// TwinCAT 3 PLC project Untitled1
// ProgramVersion: 3.1.4026.25
// libraries:
//   Tc2_Standard, * (Beckhoff Automation GmbH)
//   Tc2_System, * (Beckhoff Automation GmbH)
// project tree:
//   GVLs/ GVL_EverySignal.TcGVL, GVL_Inputs.TcGVL, GVL_IO.TcGVL, GVL_Outputs.TcGVL
//   / PlcTask.TcTTO
//   POUs/ MAIN.TcPOU, PRG_Mapping.TcPOU
// real-time tasks:
//   TASK PlcTask: cycle T#10ms, priority 20, ADS port 350
//   TASK PlcTask1: cycle T#10ms, priority 21, ADS port 351
//   TASK CNC-Task ADS: cycle default, priority 7, ADS port 558
//   TASK CNC-Task COM: cycle T#10ms, priority 14, ADS port 556
//   TASK CNC-Task SDA: cycle T#10ms, priority 9, ADS port 555
//   TASK CNC-Task GEO: cycle T#2ms, priority 3, ADS port 554
// motion (NC):
//   TASK NC-Task 1 SAF: cycle T#2ms, priority 4, ADS port 501
//   TASK NC-Task 1 SVB: cycle T#10ms, priority 8, ADS port 511
//   AXIS Axis 1 (id 1)
//     OtherSettings: AllowMotionCmdToSlave=true
//     encoder EncType=8
//       EncPara: MaxCount=#xffffffff
//     drive DrvType=9
//       DrvPara: MaxCount=#xffffffff
//         Analog: VeloScale=6, TorqueSetpointScale=10, ScaleFactorActTorque=0.1
//         TimeComp: TaskDelayCycles=1
//     controller CtrType=1
//       CtrPara: PriorControlFactor=1
//         Observer: BandWidth=20
//   AXIS Axis 2 (id 2)
//     OtherSettings: AllowMotionCmdToSlave=true
//     encoder EncType=8
//       EncPara: MaxCount=#xffffffff
//     drive DrvType=9
//       DrvPara: MaxCount=#xffffffff
//         Analog: VeloScale=6, TorqueSetpointScale=10, ScaleFactorActTorque=0.1
//         TimeComp: TaskDelayCycles=1
//     controller CtrType=1
//       CtrPara: PriorControlFactor=1
//         Observer: BandWidth=20
// I/O:
//   DEVICE C6015 (X102), AmsNetId 192.168.0.101.2.1
//     EtherCAT1  (CU1128) Junction [CU1128 6x EtherCAT junction] // Connected to PLC (C6015) using X1
//       (AX5206-0000-0011) EtherCAT4 [AX5206-0000-0011 EtherCAT Drive (SoE, 2 Ch.)] // Attached to EtherCAT1 at EtherCAT
//       EtherCAT2  (EK1100) Coupler MP-6K1 [EK1100 EtherCAT Coupler (2A E-Bus)] // Connected to EtherCAT1, Junction at X1 (W EtherCAT2 RS PRO 240-6302 1m 4x0.14 5.1)
//         (EL1809) Input Terminal MP-6K10 [EL1809 16Ch. Dig. Input 24V, 3ms] // Attached to EtherCAT 2 Coupler
//         (EL2809) Output Teminal MP-6K20 [EL2809 16Ch. Dig. Output 24V, 0.5A] // Attached to EtherCAT2 Coupler
//       Box 8 (EP1018-0001) MS-9K1 [EP1018-0001 8 Ch. Dig. Input 24V, 10µs, M8]
//       Box 9 (EP1018-0001) MS-9K2 [EP1018-0001 8 Ch. Dig. Input 24V, 10µs, M8]
//       Box 10 (EP1018-0001) MS-9K3 [EP1018-0001 8 Ch. Dig. Input 24V, 10µs, M8]
//       Box 11 (EP2028-0001) MS-10K1 [EP2028-0001 8 Ch. Dig. Output 24V, 2A, M8]
//       Box 12 (EP2028-0001) MS-10K2 [EP2028-0001 8 Ch. Dig. Output 24V, 2A, M8]
//       EtherCAT3 (EK1100) Coupler LS-7K1 [EK1100 EtherCAT Coupler (2A E-Bus)] // Attached to EtherCAT1, Junction at X1 (W EtherCAT3 RS PRO 240-6325 5m 4x0.14)
//         (EL1809) Input Terminal LS-7K10 [EL1809 16Ch. Dig. Input 24V, 3ms] // Attached to EtherCAT3 Coupler
//         (EL2809) Output Terminal LS-7K20 [EL2809 16Ch. Dig. Output 24V, 0.5A] // Attached to EtherCAT3 Coupler
//       Box 2 (CU1128-B) [CU1128 6x EtherCAT junction - Dev A]
//       Box 3 (CU1128-C) [CU1128 6x EtherCAT junction - Dev B]
// variable links:
//   Untitled1/Untitled1 Instance <-> C6015 (X102)/EtherCAT1  (CU1128) Junction/Box 10 (EP1018-0001) MS-9K3
//     PlcTask Inputs/GVL_IO.DI_E1052_{0..7} <-> Channel {1..8}/E1052.{0..7}_X{1..8}:4_DI{0..7}  (8 links)
//   Untitled1/Untitled1 Instance <-> C6015 (X102)/EtherCAT1  (CU1128) Junction/Box 11 (EP2028-0001) MS-10K1
//     PlcTask Outputs/GVL_IO.DQ_A1050_{0..7} <-> Channel {1..8}/A1050.{0..7}_X{1..8}:4_DQ{0..7}  (8 links)
//   Untitled1/Untitled1 Instance <-> C6015 (X102)/EtherCAT1  (CU1128) Junction/Box 12 (EP2028-0001) MS-10K2
//     PlcTask Outputs/GVL_IO.DQ_A1051_{0..7} <-> Channel {1..8}/A1051.{0..7}_X{1..8}:4_DQ{0..7}  (8 links)
//   Untitled1/Untitled1 Instance <-> C6015 (X102)/EtherCAT1  (CU1128) Junction/Box 8 (EP1018-0001) MS-9K1
//     PlcTask Inputs/GVL_IO.DI_E1050_0 <-> Channel 1/E1050.0 _X1:4_DI0
//     PlcTask Inputs/GVL_IO.DI_E1050_{1..5} <-> Channel {2..6}/E1050.{1..5}_X{2..6}:4_DI{1..5}  (5 links)
//   Untitled1/Untitled1 Instance <-> C6015 (X102)/EtherCAT1  (CU1128) Junction/Box 9 (EP1018-0001) MS-9K2
//     PlcTask Inputs/GVL_IO.DI_E1051_{0..3} <-> Channel {1..4}/E1051.{0..3}_X{1..4}:4_DI{0..3}  (4 links)
//   Untitled1/Untitled1 Instance <-> C6015 (X102)/EtherCAT1  (CU1128) Junction/EtherCAT2  (EK1100) Coupler MP-6K1/(EL1809) Input Terminal MP-6K10
//     PlcTask Inputs/GVL_IO.DI_E0_0 <-> Channel 1/E0.0_1_DI0
//     PlcTask Inputs/GVL_IO.DI_E0_1 <-> Channel 2/E0.1_2_DI1
//   Untitled1/Untitled1 Instance <-> C6015 (X102)/EtherCAT1  (CU1128) Junction/EtherCAT2  (EK1100) Coupler MP-6K1/(EL2809) Output Teminal MP-6K20
//     PlcTask Outputs/GVL_IO.DQ_A0_0 <-> Channel 1/A0.0_1_DQ0
//     PlcTask Outputs/GVL_IO.DQ_A0_1 <-> Channel 2/A0.1_2_DQ1
//   Untitled1/Untitled1 Instance <-> C6015 (X102)/EtherCAT1  (CU1128) Junction/EtherCAT3 (EK1100) Coupler LS-7K1/ (EL2809) Output Terminal LS-7K20
//     PlcTask Outputs/GVL_IO.DQ_A50_{0..5} <-> Channel {1..6}/A50.{0..5}_{1..6}_DQ{0..5}  (6 links)
//   Untitled1/Untitled1 Instance <-> C6015 (X102)/EtherCAT1  (CU1128) Junction/EtherCAT3 (EK1100) Coupler LS-7K1/(EL1809) Input Terminal LS-7K10
//     PlcTask Inputs/GVL_IO.DI_E50_0 <-> Channel 1/E50.0_1_DI0
//     PlcTask Inputs/GVL_IO.DI_E50_1 <-> Channel 2/E50.1_2_DI1
//     PlcTask Inputs/GVL_IO.DI_E50_2 <-> Channel 3/E50.2_3_DI2

CONFIGURATION Untitled1
    RESOURCE PLC ON TwinCAT3
        TASK PlcTask(INTERVAL := T#10ms, PRIORITY := 21);
        PROGRAM MAIN WITH PlcTask : MAIN;
    END_RESOURCE
END_CONFIGURATION

// ---- GVLs/GVL_EverySignal.TcGVL
{attribute 'qualified_only'}
VAR_GLOBAL
	//======= INPUTS ======
	
	// Safety
	bWartungseinheitDruckschalter	: BOOL;   //MaintenanceUnitPressureSwitch
	bNotHaltBetatigt				: BOOL;   //EmergencyStopActivated
	
	// CW
	bCWLReady						: BOOL;   
	bCWJobLoaded					: BOOL;
	bCWMarkInProgress				: BOOL;
	
	// Infeed
	bLichtschrankeEinlauf			: BOOL;   //InfeedLightBarrier
	bServoEinlaufEingerastet		: BOOL;   //ServoInletLockedIntoPlace
	bServoEinlaufAS					: BOOL;   //ServoInfeed
	bServoEinlaufGS					: BOOL;   //ServoInfeed
	
	// Outfeed
	bLichtschrankeAuslauf			: BOOL;   //OutfeedLightBarrier
	bServoAuslaufEingerastet		: BOOL;   //ServoOutletLockedIntoPlace
	bServoAuslaufAS					: BOOL;   //ServoOutlet
	bServoAuslaufGS					: BOOL;   //ServoOutlet
	
	// Ejector
	bZylinderAuswerfwerAS			: BOOL;   //CylinderEjector
	bZylinderAuswerferGS			: BOOL;   //CylinderEjector
	
	// Clamp
	bZylinderSpannerAS				: BOOL;   //CylinderClamp
	bZylinderSpannerGS				: BOOL;   //CylinderClamp
	
	// Diverter
	bZylinderWeicheAS				: BOOL;   //CylinderDiverter
	bZylinderWeicheGS				: BOOL;   //CylinderDiverter
	
	
	
	
	//======== OUTPUTS ========
	
	//Valve
	bVentilAuswerferAS				: BOOL;   //ValveEjector
	bVentilAuswerferGS				: BOOL;   //ValveEjector
	
	bVentilSpannerAS				: BOOL;   //ValveClamp
	bVentilSpannerGS				: BOOL;   //ValveClamp
	
	bVentilWeicheAS					: BOOL;   //ValveDiverter
	bVentilWeicheGS					: BOOL;   //ValveDiverter
	
	bVentilAusblastenAS				: BOOL;   //BlowOutValve
	bVentilAusblastenGS				: BOOL;   //BlowOutValve
	
	bVentilEinlaufAS				: BOOL;   //ValveInfeed
	bVentilEinlaufGS				: BOOL;   //ValveInfeed
	
	bVentilAuslaufAS				: BOOL;   //ValveOutfeed
	bVentilAuslaufGS				: BOOL;   //ValveOutfeed
	
	bVentilAuswerfBypassAS			: BOOL;   //EjectionBypassValve
	bVentilAuswerfBypassGS			: BOOL;   //EjectionBypassValve
	
	// CW
	bCWTrigger						: BOOL;
	bCWSTO							: BOOL;
	bJob							: BOOL;
	
	// Machine
	bWartungseinheitEntluften		: BOOL;   //MaintenanceUnitVenting
	bLaserEnable					: BOOL;

END_VAR

// ---- GVLs/GVL_Inputs.TcGVL
{attribute 'qualified_only'}
VAR_GLOBAL
	bWartungseinheitDruckschalter	: BOOL;   //MaintenanceUnitPressureSwitch
	bNotHaltBetatigt				: BOOL;   //EmergencyStopActivated
	
	bCWLReady						: BOOL;   
	bCWJobLoaded					: BOOL;
	bCWMarkInProgress				: BOOL;
	
	bZylinderAuswerferAS			: BOOL;   //CylinderEjector
	bZylinderAuswerferGS			: BOOL;   //CylinderEjector
	bZylinderSpannerAS				: BOOL;   //CylinderClamp
	bZylinderSpannerGS				: BOOL;   //CylinderClamp
	bZylinderWeicheAS				: BOOL;   //CylinderDiverter
	bZylinderWeicheGS				: BOOL;   //CylinderDiverter
	
	bZylinderEinlaufAS				: BOOL;	  //CylinderInfeed
	bZylinderEinlaufGS				: BOOL;	  //CylinderInfeed
	bZylinderAuslaufAS				: BOOL;	  //CylinderOutfeed
	bZylinderAuslaufGS				: BOOL;	  //CylinderOutfeed
	
	bLichtschrankeEinlauf			: BOOL;   //InfeedLightBarrier
	bServoEinlaufEingerastet		: BOOL;   //ServoInletLockedIntoPlace
	bServoEinlaufAS					: BOOL;   //ServoInfeed
	bServoEinlaufGS					: BOOL;   //ServoInfeed
	bLichtschrankeAuslauf			: BOOL;   //OutfeedLightBarrier
	bServoAuslaufEingerastet		: BOOL;   //ServoOutletLockedIntoPlace
	bServoAuslaufAS					: BOOL;   //ServoOutlet
	bServoAuslaufGS					: BOOL;   //ServoOutlet
	
		

END_VAR

// ---- GVLs/GVL_IO.TcGVL
{attribute 'qualified_only'}
VAR_GLOBAL
	//Inputs
	DI_E0_0     AT%I*	:BOOL;
	DI_E0_1		AT%I*	:BOOL;
	
	DI_E50_0	AT%I*	:BOOL;
	DI_E50_1	AT%I*	:BOOL;
	DI_E50_2	AT%I*	:BOOL;
	
	DI_E1050_0	AT%I*	:BOOL;
	DI_E1050_1	AT%I*	:BOOL;
	DI_E1050_2	AT%I*	:BOOL;
	DI_E1050_3	AT%I*	:BOOL;
	DI_E1050_4	AT%I*	:BOOL;
	DI_E1050_5	AT%I*	:BOOL;
	
	DI_E1051_0	AT%I*	:BOOL;
	DI_E1051_1	AT%I*	:BOOL;
	DI_E1051_2	AT%I*	:BOOL;
	DI_E1051_3	AT%I*	:BOOL;
	
	DI_E1052_0	AT%I*	:BOOL;
	DI_E1052_1	AT%I*	:BOOL;
	DI_E1052_2	AT%I*	:BOOL;
	DI_E1052_3	AT%I*	:BOOL;
	DI_E1052_4	AT%I*	:BOOL;
	DI_E1052_5	AT%I*	:BOOL;
	DI_E1052_6	AT%I*	:BOOL;
	DI_E1052_7	AT%I*	:BOOL;
	
	
	//Outputs
	DQ_A0_0		AT%Q*	:BOOL;
	DQ_A0_1		AT%Q*	:BOOL;
	
	DQ_A50_0	AT%Q*	:BOOL;
	DQ_A50_1	AT%Q*	:BOOL;
	DQ_A50_2	AT%Q*	:BOOL;
	DQ_A50_3	AT%Q*	:BOOL;
	DQ_A50_4	AT%Q*	:BOOL;
	DQ_A50_5	AT%Q*	:BOOL;
	
	DQ_A1050_0	AT%Q*	:BOOL;
	DQ_A1050_1	AT%Q*	:BOOL;
	DQ_A1050_2	AT%Q*	:BOOL;
	DQ_A1050_3	AT%Q*	:BOOL;
	DQ_A1050_4	AT%Q*	:BOOL;
	DQ_A1050_5	AT%Q*	:BOOL;
	DQ_A1050_6	AT%Q*	:BOOL;
	DQ_A1050_7	AT%Q*	:BOOL;
	
	DQ_A1051_0	AT%Q*	:BOOL;
	DQ_A1051_1	AT%Q*	:BOOL;
	DQ_A1051_2	AT%Q*	:BOOL;
	DQ_A1051_3	AT%Q*	:BOOL;
	DQ_A1051_4	AT%Q*	:BOOL;
	DQ_A1051_5	AT%Q*	:BOOL;
	DQ_A1051_6	AT%Q*	:BOOL;
	DQ_A1051_7	AT%Q*	:BOOL;
	
	
END_VAR

// ---- GVLs/GVL_Outputs.TcGVL
{attribute 'qualified_only'}
VAR_GLOBAL
	bWartungseinheitEntluften		: BOOL;   //MaintenanceUnitVenting
	bLaserEnable					: BOOL;

	bCWTrigger						: BOOL;
	bCWSTO							: BOOL;
	bCWJob							: BOOL;

	bVentilAuswerferAS				: BOOL;   //ValveEjector
	bVentilAuswerferGS				: BOOL;   //ValveEjector
	bVentilSpannerAS				: BOOL;   //ValveClamp
	bVentilSpannerGS				: BOOL;   //ValveClamp
	bVentilWeicheAS					: BOOL;   //ValveDiverter
	bVentilWeicheGS					: BOOL;   //ValveDiverter
	bVentilAusblastenAS				: BOOL;   //BlowOutValve
	bVentilAusblastenGS				: BOOL;   //BlowOutValve	
	
	bVentilEinlaufAS				: BOOL;   //ValveInfeed
	bVentilEinlaufGS				: BOOL;   //ValveInfeed
	bVentilAuslaufAS				: BOOL;   //ValveOutfeed
	bVentilAuslaufGS				: BOOL;   //ValveOutfeed	
	bVentilAuswerfBypassAS			: BOOL;   //EjectionBypassValve
	bVentilAuswerfBypassGS			: BOOL;   //EjectionBypassValve

END_VAR

// ---- POUs/MAIN.TcPOU
PROGRAM MAIN
VAR
END_VAR

END_PROGRAM

// ---- POUs/PRG_Mapping.TcPOU
PROGRAM PRG_Mapping
VAR
END_VAR

//=== Mapping the input signals

GVL_Inputs.bWartungseinheitDruckschalter := GVL_IO.DI_E0_0;
GVL_Inputs.bNotHaltBetatigt := GVL_IO.DI_E0_1;

GVL_Inputs.bCWLReady := GVL_IO.DI_E50_0;
GVL_Inputs.bCWJobLoaded := GVL_IO.DI_E50_1;
GVL_Inputs.bCWMarkInProgress := GVL_IO.DI_E50_2;

GVL_Inputs.bZylinderAuswerferAS := GVL_IO.DI_E1050_0;
GVL_Inputs.bZylinderAuswerferGS := GVL_IO.DI_E1050_1;
GVL_Inputs.bZylinderSpannerAS := GVL_IO.DI_E1050_2;
GVL_Inputs.bZylinderSpannerGS := GVL_IO.DI_E1050_3;
GVL_Inputs.bZylinderWeicheAS := GVL_IO.DI_E1050_4;
GVL_Inputs.bZylinderWeicheGS := GVL_IO.DI_E1050_5;

GVL_Inputs.bZylinderEinlaufAS := GVL_IO.DI_E1051_0;
GVL_Inputs.bZylinderEinlaufGS := GVL_IO.DI_E1051_1;
GVL_Inputs.bZylinderAuslaufAS := GVL_IO.DI_E1051_2;
GVL_Inputs.bZylinderAuslaufGS := GVL_IO.DI_E1051_3;

GVL_Inputs.bLichtschrankeEinlauf := GVL_IO.DI_E1052_0;
GVL_Inputs.bServoEinlaufEingerastet := GVL_IO.DI_E1052_1;
GVL_Inputs.bServoEinlaufAS := GVL_IO.DI_E1052_2;
GVL_Inputs.bServoEinlaufGS := GVL_IO.DI_E1052_3;
GVL_Inputs.bLichtschrankeAuslauf := GVL_IO.DI_E1052_4;
GVL_Inputs.bServoAuslaufEingerastet := GVL_IO.DI_E1052_5;
GVL_Inputs.bServoAuslaufAS := GVL_IO.DI_E1052_6;
GVL_Inputs.bServoAuslaufGS := GVL_IO.DI_E1052_7;


//=== Mapping the output signals

GVL_Outputs.bWartungseinheitEntluften := GVL_IO.DQ_A0_0;
GVL_Outputs.bLaserEnable := GVL_IO.DQ_A0_1;

GVL_Outputs.bCWTrigger := GVL_IO.DQ_A50_0;
GVL_Outputs.bCWJob := GVL_IO.DQ_A50_1;
GVL_Outputs.bCWJob := GVL_IO.DQ_A50_2;
GVL_Outputs.bCWJob := GVL_IO.DQ_A50_3;
GVL_Outputs.bCWJob := GVL_IO.DQ_A50_4;
GVL_Outputs.bCWSTO := GVL_IO.DQ_A50_5;

GVL_Outputs.bVentilAuswerferAS := GVL_IO.DQ_A1050_0;
GVL_Outputs.bVentilAuswerferGS := GVL_IO.DQ_A1050_1;
GVL_Outputs.bVentilSpannerAS := GVL_IO.DQ_A1050_2;
GVL_Outputs.bVentilSpannerGS := GVL_IO.DQ_A1050_3;
GVL_Outputs.bVentilWeicheAS := GVL_IO.DQ_A1050_4;
GVL_Outputs.bVentilWeicheGS := GVL_IO.DQ_A1050_5;
GVL_Outputs.bVentilAusblastenAS := GVL_IO.DQ_A1050_6;
GVL_Outputs.bVentilAusblastenGS := GVL_IO.DQ_A1050_7;

GVL_Outputs.bVentilEinlaufAS := GVL_IO.DQ_A1051_0;
GVL_Outputs.bVentilEinlaufGS := GVL_IO.DQ_A1051_1;
GVL_Outputs.bVentilAuslaufAS := GVL_IO.DQ_A1051_2;
GVL_Outputs.bVentilAuslaufGS := GVL_IO.DQ_A1051_3;
GVL_Outputs.bVentilAusblastenAS := GVL_IO.DQ_A1051_4;
GVL_Outputs.bVentilAusblastenGS := GVL_IO.DQ_A1051_5;
GVL_Outputs.bVentilAuswerfBypassAS := GVL_IO.DQ_A1051_6;
GVL_Outputs.bVentilAuswerfBypassGS := GVL_IO.DQ_A1051_7;

END_PROGRAM
